Fanuc KAREL source: ko00046.KL

-- PROVISIONAL review KL for V1013-1; original PC SHA256 61799707e98ebbcb1868e0261da0690aeec2e9e569baa7e2baee15e7db781f4e
-- Incomplete behavior may be omitted. Consult companion uncertainty JSON. Do not deploy.
PROGRAM KO00046
%NOLOCKGROUP
BEGIN
  -- UNRESOLVED_PC offsets 5-12; opcodes 9D,23
  -- UNRESOLVED_PC offsets 17-69; opcodes 27,27,49,7E,AD,27,49,7E,AD,22,31,7E,4A
  -- UNRESOLVED_PC offsets 74-78; opcodes 7F
END KO00046
